FUNCTION_BLOCK FB_PI_Controller_Tests EXTENDS TcUnit.FB_TestSuite

Test_ProportionalOnlyWithBias();
Test_OutputClampedToMax();
Test_OutputClampedToMin();
Test_IntegralInRepeatsPerMinute();
Test_IntegralInRepeatsPerSecond();
Test_UsesCycleTimeOfCallingTask();

METHOD PRIVATE Test_ProportionalOnlyWithBias
VAR
  pi : FB_PI_Controller;
END_VAR
TcUnit.TEST(__POUNAME());

pi(ProcessVariable := 4.0, Setpoint := 10.0, Kp := 2.0, IntegralConstant := 0.0, MaxLoopOutput := 100.0, MinLoopOutput := -100.0, Bias := 1.0);
AssertEquals_LREAL(Expected := 13.0, Actual := pi.Output, Delta := 1.0E-9, Message := 'Kp * error + bias');

TEST_FINISHED_NAMED(__POUNAME());
END_METHOD

METHOD PRIVATE Test_OutputClampedToMax
VAR
  pi : FB_PI_Controller;
END_VAR
TcUnit.TEST(__POUNAME());

pi(ProcessVariable := 4.0, Setpoint := 10.0, Kp := 2.0, IntegralConstant := 0.0, MaxLoopOutput := 5.0, MinLoopOutput := -100.0, Bias := 0.0);
AssertEquals_LREAL(Expected := 5.0, Actual := pi.Output, Delta := 1.0E-9, Message := 'output held at the maximum');

TEST_FINISHED_NAMED(__POUNAME());
END_METHOD

METHOD PRIVATE Test_OutputClampedToMin
VAR
  pi : FB_PI_Controller;
END_VAR
TcUnit.TEST(__POUNAME());

pi(ProcessVariable := 10.0, Setpoint := 4.0, Kp := 2.0, IntegralConstant := 0.0, MaxLoopOutput := 100.0, MinLoopOutput := -5.0, Bias := 0.0);
AssertEquals_LREAL(Expected := -5.0, Actual := pi.Output, Delta := 1.0E-9, Message := 'output held at the minimum');

TEST_FINISHED_NAMED(__POUNAME());
END_METHOD

METHOD PRIVATE Test_IntegralInRepeatsPerMinute
VAR
  pi : FB_PI_Controller;
END_VAR
TcUnit.TEST(__POUNAME());

// 60 repeats per minute is 1 repeat per second: one 10 ms cycle adds error * 0.01
pi(ProcessVariable := 0.0, Setpoint := 1.0, Kp := 0.0, IntegralConstant := 60.0, RepeatsPerMinute := TRUE, MaxLoopOutput := 100.0, MinLoopOutput := -100.0, Bias := 0.0);
AssertEquals_LREAL(Expected := 0.01, Actual := pi.Output, Delta := 1.0E-6, Message := 'integral normalised from repeats per minute');

TEST_FINISHED_NAMED(__POUNAME());
END_METHOD

METHOD PRIVATE Test_IntegralInRepeatsPerSecond
VAR
  pi : FB_PI_Controller;
END_VAR
TcUnit.TEST(__POUNAME());

pi(ProcessVariable := 0.0, Setpoint := 1.0, Kp := 0.0, IntegralConstant := 1.0, RepeatsPerMinute := FALSE, MaxLoopOutput := 100.0, MinLoopOutput := -100.0, Bias := 0.0);
AssertEquals_LREAL(Expected := 0.01, Actual := pi.Output, Delta := 1.0E-6, Message := 'integral in repeats per second');

TEST_FINISHED_NAMED(__POUNAME());
END_METHOD

METHOD PRIVATE Test_UsesCycleTimeOfCallingTask
TcUnit.TEST(__POUNAME());

IF NOT ControllersInSlowTask.HasRunOnce THEN
  RETURN;
END_IF

AssertEquals_LREAL(Expected := 0.05, Actual := ControllersInSlowTask.PiOutput, Delta := 1.0E-6, Message := 'one cycle of the 50 ms SlowTask, not the 10 ms PlcTask');

TEST_FINISHED_NAMED(__POUNAME());
END_METHOD

END_FUNCTION_BLOCK

(* stored: Version 1.1.0.1, ProductVersion 3.1.4026.22
   POU FB_PI_Controller_Tests: Id {64e85ef2-1068-4d81-9e39-ee7c784040f8}, SpecialFunc None
   Method Test_ProportionalOnlyWithBias: Id {cd21461c-a771-480f-9b38-caf06491bc0a}
   Method Test_OutputClampedToMax: Id {b33ce352-b16b-4762-acc8-ec222d717a77}
   Method Test_OutputClampedToMin: Id {531a44cf-2575-4534-80f4-5228eaefdb1f}
   Method Test_IntegralInRepeatsPerMinute: Id {adebae75-f62e-4eb2-b21c-bb273750d426}
   Method Test_IntegralInRepeatsPerSecond: Id {4b355492-b074-4b29-a973-191979cb2e91}
   Method Test_UsesCycleTimeOfCallingTask: Id {7f10557a-0361-4a01-b733-27f389d6ed94} *)
